FUNCTION_BLOCK FB_1001_Station1
VAR_INPUT
    i_bEnable : BOOL;
END_VAR
VAR_OUTPUT
    q_bDone : BOOL;
END_VAR
BEGIN
    ;
END_FUNCTION_BLOCK
